(* IEC 61131-3 sources: Zbiorniki_user/Temp/Import/MpRecipe, 4 files *)

(* ---- MpRecipe.typ ---- *)
TYPE
	MpRecipeStatusIDType : 	STRUCT
		ID : MpRecipeErrorEnum; (*Error code for mapp component*)
		Severity : MpComSeveritiesEnum; (*Describes the type of information supplied by the status ID (success, information, warning, error)*)
		Code : UINT; (*Code for the status ID. This error number can be used to search for additional information in the help system*)
	END_STRUCT;
	MpRecipeDiagType : 	STRUCT
		StatusID : MpRecipeStatusIDType; (*StatusID diagnostics structure*)
	END_STRUCT;
	MpRecipeInfoType : 	STRUCT
		Diag : MpRecipeDiagType; (*Diagnostic structure for the status ID*)
	END_STRUCT;
	MpRecipeUISetupConfirmType : 	STRUCT
		RecipeLoad : BOOL; (*Enables a confirmation window when loading a recipe*)
		RecipeSave : BOOL; (*Enables a confirmation window when saving a recipe*)
		RecipeCreate : BOOL; (*Enables a confirmation window when creating a recipe	*)
		RecipeDelete : BOOL; (*Enables a confirmation window when creating a recipe*)
		RecipeRename : BOOL; (*Enables a confirmation window when renaming a recipe*)
	END_STRUCT;
	MpRecipeUISetupType : 	STRUCT
		RecipeListSize : UINT := 20; (*Number of recipes to be displayed on one page of the list in the HMI application*)
		RecipeListScrollWindow : USINT := 1; (*Determines how many entries from the list are displayed in advance when scrolling up and down*)
		Confirmation : MpRecipeUISetupConfirmType; (*Displaying the confirmation window*)
		AutoLoadHeader : BOOL; (*Header info of a recipe should be loaded automatically when a recipe is selected (like a preview) *)
	END_STRUCT;
	MpRecipeUIMessageEnum :
		(
		mpRECIPE_UI_MSG_NONE := 0, (*No dialog is required*)
		mpRECIPE_UI_MSG_CONFIRM_LOAD := 1, (*Dialog box for confirming the loading procedure*)
		mpRECIPE_UI_MSG_CONFIRM_SAVE := 2, (*Dialog box for confirming the saving procedure*)
		mpRECIPE_UI_MSG_CONFIRM_CREATE := 3, (*Dialog box for confirming the creation of a new recipe	*)
		mpRECIPE_UI_MSG_CONFIRM_DELETE := 4, (*Dialog box for confirming the deletion of an existing recipe*)
		mpRECIPE_UI_MSG_CONFIRM_RENAME := 5 (*Dialog box for confirming the renaming of an existing recipe*)
		);
	MpRecipeUIStatusEnum :
		(
		mpRECIPE_UI_STATUS_IDLE := 0, (*Indicates that no process is currently active*)
		mpRECIPE_UI_STATUS_LOAD := 1, (*A recipe is being loaded*)
		mpRECIPE_UI_STATUS_SAVE := 2, (*A recipe is being saved*)
		mpRECIPE_UI_STATUS_CREATE := 3, (*A recipe is being created*)
		mpRECIPE_UI_STATUS_REFRESH := 4, (*The recipe list is being refreshed*)
		mpRECIPE_UI_STATUS_NOTIFY := 5, (*mapp components are being informed that new parameters are to be used*)
		mpRECIPE_UI_STATUS_DELETE := 6, (*A recipe is being deleted*)
		mpRECIPE_UI_STATUS_RENAME := 7, (*A recipe is being renamed*)
		mpRECIPE_UI_STATUS_ERROR := 99 (*The last operation generated an error*)
		);
	MpRecipeUIMessageBoxType : 	STRUCT
		LayerStatus : UINT; (*Visibility of the dialog box *)
		Type : MpRecipeUIMessageEnum; (*Type of dialog box*)
		Confirm : BOOL; (*Confirms the operation*)
		Cancel : BOOL; (*Cancels the operation*)
	END_STRUCT;
	MpRecipeUINewType : 	STRUCT
		FileName : STRING[255]; (*Name of the new recipe*)
		Create : BOOL; (*Creates a new recipe*)
	END_STRUCT;
	MpRecipeUIConnectType : 	STRUCT
		Status : MpRecipeUIStatusEnum; (*Current operation*)
		Recipe : MpRecipeUIRecipeType; (*Access to existing recipes*)
		New : MpRecipeUINewType; (*To create new recipes*)
		MessageBox : MpRecipeUIMessageBoxType; (*Controls dialog boxes*)
		DefaultLayerStatus : UINT; (*Status data point for the default layer of the visualization page where the recipe management system is being displayed*)
	END_STRUCT;
	MpRecipeUIRecipeListType : 	STRUCT
		Names : ARRAY[0..19] OF STRING[255]; (*List of all available recipes (filenames)*)
		SelectedIndex : UINT; (*Index of the entry currently selected in the list*)
		MaxSelection : UINT; (*Index of the last entry in the list*)
		PageUp : BOOL; (*Jumps to the start of the current page and then scrolls up one page at a time *)
		PageDown : BOOL; (*Jumps to the end of the current page and then scrolls down one page at a time *)
		StepUp : BOOL; (*Selects the previous entry in the list*)
		StepDown : BOOL; (*Selects the next entry in the list*)
		RangeStart : REAL; (*Shows a bar indicating which part of the list is currently being displayed-Start [%]*)
		RangeEnd : REAL; (*Shows a bar indicating which part of the list is currently being displayed-End [%]*)
		Sizes : ARRAY[0..19]OF UDINT; (*List of all recipe file sizes*)
		LastModified : ARRAY[0..19]OF STRING[50]; (*List of the last modification dates for all recipe files*)
	END_STRUCT;
	MpRecipeUIHeaderType : 	STRUCT
		Name : STRING[100]; (*Name of the recipe*)
		Description : STRING[255]; (*Comment that describes the recipe*)
		Version : STRING[20]; (*Version of the recipe*)
		DateTime : DATE_AND_TIME; (*Date and time the recipe was created*)
	END_STRUCT;
	MpRecipeUIRecipeType : 	STRUCT
		List : MpRecipeUIRecipeListType; (*List of all available recipes (filenames)*)
		Load : BOOL; (*Loads the selected recipe*)
		Save : BOOL; (*Saves the selected recipe*)
		Filter : STRING[255]; (*Filter used to sort the recipes*)
		SortOrder : MpRecipeUISortOrderEnum; (*Sorts the recipe list*)
		Refresh : BOOL; (*Updates the recipe list*)
		UpdateNotification : BOOL; (*Request to all mapp components to enter the current values of the recipe parameters*)
		Delete : BOOL; (*Deletes the selected recipe*)
		Rename : BOOL; (*Renames the currently selected recipe*)
		NewFileName : STRING[255]; (*Name of the new recipe*)
		Header : MpRecipeUIHeaderType; (*The header info of the currently selected recipe (is only loaded if the option is enabled in UISetup)*)
	END_STRUCT;
	MpRecipeXmlInfoType : 	STRUCT
		FileSize : UDINT; (*Size of the recipe stored on the respective data storage medium*)
		PendingSync : UDINT; (*Number of pending save notifications ("SaveNotification") that have not yet been confirmed*)
		Diag : MpRecipeDiagType; (*Diagnostic structure for the status ID *)
		LastLoadedRecipe : STRING[255]; (*The name of the last loaded recipe*)
	END_STRUCT;
	MpRecipeUISortOrderEnum :
		(
		mpRECIPE_UI_SORT_ASCENDING := 0, (*Sorts in ascending (alphabetic) order*)
		mpRECIPE_UI_SORT_DESCENDING := 1, (*Sorts in descending (alphabetic) order*)
		mpRECIPE_UI_SORT_DATE_ASCENDING := 2, (*Sorts in ascending (date/time) order*)
		mpRECIPE_UI_SORT_DATE_DESCENDING := 3 (*Sorts in descending (date/time) order*)
		);
	MpRecipeXmlHeaderType : 	STRUCT
		Name : STRING[100]; (*Name of the recipe*)
		Description : STRING[255]; (*Comment that describes the recipe*)
		Version : STRING[20]; (*Version of the recipe*)
		DateTime : DATE_AND_TIME; (*Date and time the recipe was created*)
	END_STRUCT;
	MpRecipeXmlLoadEnum :
		(
		mpRECIPE_XML_LOAD_ALL := 0, (*Loads the entire content of the recipe*)
		mpRECIPE_XML_LOAD_HEADER := 1 (*Loads only the recipe's header*)
		);
	MpRecipeCsvHeaderType : 	STRUCT
		Name : STRING[100]; (*Name of the recipe*)
		Description : STRING[255]; (*Comment that describes the recipe*)
		Version : STRING[20]; (*Version of the recipe*)
		DateTime : DATE_AND_TIME; (*Date and time the recipe was created*)
	END_STRUCT;
	MpRecipeCsvInfoType : 	STRUCT
		FileSize : UDINT; (*Size of the recipe stored on the respective data storage medium*)
		PendingSync : UDINT; (*Number of pending save notifications ("SaveNotification") that have not yet been confirmed*)
		LastLoadedRecipe : STRING[255]; (*The name of the last loaded recipe*)
		Diag : MpRecipeDiagType; (*Diagnostic structure for the status ID *)
	END_STRUCT;
	MpRecipeCsvLoadEnum :
		(
		mpRECIPE_CSV_LOAD_ALL := 0, (*Loads the entire content of the recipe*)
		mpRECIPE_CSV_LOAD_HEADER := 1 (*Loads only the recipe's header*)
		);
END_TYPE

(* ---- MpRecipeAlarm.typ ---- *)
TYPE
    MpRecipeXmlAlarmEnum :
        ( (* Alarms of MpRecipe Xml *)
        mpRECIPE_ALM_SAVE_FAILED := 0, (* Saving of recipe failed. *)
        mpRECIPE_ALM_SAVE_FAILED_PART := 1, (* Saving of recipe failed partially. Parts of the recipe could be saved. *)
        mpRECIPE_ALM_LOAD_FAILED := 2, (* Loading of recipe failed. *)
        mpRECIPE_ALM_LOAD_FAILED_PART := 3 (* Loading of recipe failed partially. Parts of the recipe could be loaded. *)
    );
END_TYPE

(* ---- MpRecipeError.typ ---- *)
TYPE
    MpRecipeErrorEnum :
        ( (* Error numbers of library MpRecipe *)
        mpRECIPE_NO_ERROR := 0, (* No error *)
        mpRECIPE_ERR_ACTIVATION := -1064239103, (* Could not create component [Error: 1, 0xc0910001] *)
        mpRECIPE_ERR_MPLINK_NULL := -1064239102, (* MpLink is NULL pointer [Error: 2, 0xc0910002] *)
        mpRECIPE_ERR_MPLINK_INVALID := -1064239101, (* MpLink connection not allowed [Error: 3, 0xc0910003] *)
        mpRECIPE_ERR_MPLINK_CHANGED := -1064239100, (* MpLink modified [Error: 4, 0xc0910004] *)
        mpRECIPE_ERR_MPLINK_CORRUPT := -1064239099, (* Invalid MpLink contents [Error: 5, 0xc0910005] *)
        mpRECIPE_ERR_MPLINK_IN_USE := -1064239098, (* MpLink already in use [Error: 6, 0xc0910006] *)
        mpRECIPE_ERR_CONFIG_INVALID := -1064239091, (* Invalid Configuration [Error: 13, 0xc091000d] *)
        mpRECIPE_ERR_SAVE_DATA := -1064140799, (* Failed to create recipe file {2:File} using device {3:Device} (Error cause: {1:ErrorNumber}) [Error: 32769, 0xc0928001] *)
        mpRECIPE_ERR_LOAD_DATA := -1064140798, (* Failed to load recipe from {2:File} using device {3:Device} (Error cause: {1:ErrorNumber}) [Error: 32770, 0xc0928002] *)
        mpRECIPE_ERR_INVALID_FILE_DEV := -1064140797, (* Invalid file device [Error: 32771, 0xc0928003] *)
        mpRECIPE_ERR_INVALID_FILE_NAME := -1064140796, (* Invalid filename [Error: 32772, 0xc0928004] *)
        mpRECIPE_ERR_CMD_IN_PROGRESS := -1064140795, (* Component currently executing command [Error: 32773, 0xc0928005] *)
        mpRECIPE_WRN_SAVE_WITH_WARN := -2137882618, (* Warnings while saving recipe [Warning: 32774, 0x80928006] *)
        mpRECIPE_WRN_LOAD_WITH_WARN := -2137882617, (* Warnings while loading recipe [Warning: 32775, 0x80928007] *)
        mpRECIPE_ERR_SAVE_WITH_ERRORS := -1064140792, (* Failed to write to recipe file {2:File} (Error cause: {1:ErrorNumber}) [Error: 32776, 0xc0928008] *)
        mpRECIPE_ERR_LOAD_WITH_ERRORS := -1064140791, (* Error converting recipe to parameters [Error: 32777, 0xc0928009] *)
        mpRECIPE_ERR_MISSING_RECIPE := -1064140790, (* No connection to parent component [Error: 32778, 0xc092800a] *)
        mpRECIPE_ERR_MISSING_MPFILE := -1064140789, (* No connection to file manager [Error: 32779, 0xc092800b] *)
        mpRECIPE_ERR_INVALID_SORT_ORDER := -1064140788, (* Invalid sort order selected [Error: 32780, 0xc092800c] *)
        mpRECIPE_WRN_MISSING_UICONNECT := -2137882611, (* Invalid value for "UIConnect" [Warning: 32781, 0x8092800d] *)
        mpRECIPE_ERR_INVALID_PV_NAME := -1064140786, (* Invalid PV [Error: 32782, 0xc092800e] *)
        mpRECIPE_ERR_INVALID_LOAD_TYPE := -1064140785, (* Invalid LoadType [Error: 32783, 0xc092800f] *)
        mpRECIPE_ERR_LISTING_FILES := -1064140784, (* Error creating file list [Error: 32784, 0xc0928010] *)
        mpRECIPE_ERR_PV_NAME_NULL := -1064140783, (* PV name is NULL [Error: 32785, 0xc0928011] *)
        mpRECIPE_WRN_NO_PV_REGISTERED := -2137882606, (* No PV registered [Warning: 32786, 0x80928012] *)
        mpRECIPE_ERR_SYNC_SAVE_ACTIVE := -1064140781, (* Saving active [Error: 32787, 0xc0928013] *)
        mpRECIPE_ERR_DELETING_FILE := -1064140780, (* Failed to delete recipe {2:Recipe} from device {3:Device} (Error cause: {1:ErrorNumber}) [Error: 32788, 0xc0928014] *)
        mpRECIPE_WRN_EMPTY_RECIPE := -2137882603, (* Saving empty recipe file [Warning: 32789, 0x80928015] *)
        mpRECIPE_INF_WAIT_RECIPE_FB := 1083342870, (* Waiting for parent recipe component [Informational: 32790, 0x40928016] *)
        mpRECIPE_ERR_RENAMING_FILE := -1064140777, (* Failed to rename recipe {2:FromName} to {3:ToName} (Error cause: {1:ErrorNumber} [Error: 32791, 0xc0928017] *)
        mpRECIPE_WRN_NO_PV_FOUND := -2137882600, (* None of the registered PVs were found in the recipe file while loading. The file might be corrupted. [Warning: 32792, 0x80928018] *)
        mpRECIPE_WRN_LIST_SIZE := -2137882599 (* The UISetup.RecipeListSize {2:Size} is out of limit (1-20). [Warning: 32793, 0x80928019] *)
        );
END_TYPE

(* ---- MpRecipe.fun ---- *)
FUNCTION_BLOCK MpRecipeRegParSync (*Declare a PV as a recipe parameter and perform synchronisation*) (* $GROUP=mapp Services,$CAT=XML Recipe,$GROUPICON=Icon_mapp.png,$CATICON=Icon_MpRecipe.png *)
	VAR_INPUT
		MpLink : REFERENCE TO MpComIdentType; (*Connection to mapp*) (* *) (*#PAR#;*)
		Enable : BOOL; (*Enables/Disables the function block *) (* *) (*#PAR#;*)
		ErrorReset : BOOL; (*Resets function block errors*) (* *) (*#PAR#;*)
		PVName : REFERENCE TO STRING[100]; (*Name of the PV that should be saved to the recipe*) (* *) (*#PAR#;*)
		Category : REFERENCE TO STRING[50]; (*Name of the category used to organize the parameters*) (* *) (*#PAR#OPT#;*)
		ConfirmSave : BOOL; (*Confirms that the current data of the registered PV can be saved to the recipe. This is used in connection with "SaveNotification"*) (* *) (*#CMD#;*)
	END_VAR
	VAR_OUTPUT
		Active : BOOL; (*Indicates whether the function block is active*) (* *) (*#PAR#;*)
		Error : BOOL; (*Indicates that the function block is in an error state or a command was not executed correctly*) (* *) (*#PAR#;*)
		StatusID : DINT; (*Status information about the function block*) (* *) (*#PAR#; *)
		UpdateNotification : BOOL; (*TRUE if a new recipe has been loaded and the registered PV contains new values. This is automatically reset after one cycle*) (* *) (*#CMD#OPT#;*)
		SaveNotification : BOOL; (*TRUE if a recipe is saved and new data should be copied to the recipe, but before the data is actually transferred to the recipe. This is used in connection with "ConfirmSave"*) (* *) (*#CMD#;*)
		Info : MpRecipeInfoType; (*Additional information about the component*) (* *) (*#CMD#;*)
	END_VAR
	VAR
		Internal : {REDUND_UNREPLICABLE} MpComInternalDataType; (*Internal stucture*) (* *) (*#OMIT#;*)
	END_VAR
END_FUNCTION_BLOCK

FUNCTION_BLOCK MpRecipeRegPar (*Declare a PV as a recipe parameter*) (* $GROUP=mapp Services,$CAT=XML Recipe,$GROUPICON=Icon_mapp.png,$CATICON=Icon_MpRecipe.png *)
	VAR_INPUT
		MpLink : REFERENCE TO MpComIdentType; (* Connection to mapp*) (* *) (*#PAR#;*)
		Enable : BOOL; (*Enables/Disables the function block*) (* *) (*#PAR#;*)
		ErrorReset : BOOL; (*Resets function block errors*) (* *) (*#PAR#;*)
		PVName : REFERENCE TO STRING[100]; (*Name of the PV that should be saved to the recipe*) (* *) (*#PAR#;*)
		Category : REFERENCE TO STRING[50]; (*Name of the category used to organize the parameters*) (* *) (*#PAR#OPT#;*)
	END_VAR
	VAR_OUTPUT
		Active : BOOL; (*Indicates whether the function block is active*) (* *) (*#PAR#;*)
		Error : BOOL; (*Indicates that the function block is in an error state or a command was not executed correctly*) (* *) (*#PAR#;*)
		StatusID : DINT; (*Status information about the function block*) (* *) (*#PAR#; *)
		UpdateNotification : BOOL; (*TRUE if a new recipe has been loaded and the registered PV contains new values. This is automatically reset after one cycle*) (* *) (*#CMD#OPT#;*)
		Info : MpRecipeInfoType; (*Additional information about the component*) (* *) (*#CMD#;*)
	END_VAR
	VAR
		Internal : {REDUND_UNREPLICABLE} MpComInternalDataType; (*Internal stucture*) (* *) (*#OMIT#;*)
	END_VAR
END_FUNCTION_BLOCK

FUNCTION_BLOCK MpRecipeXml (*Load/save parameters from/to an XML file*) (* $GROUP=mapp Services,$CAT=XML Recipe,$GROUPICON=Icon_mapp.png,$CATICON=Icon_MpRecipe.png *)
	VAR_INPUT
		MpLink : REFERENCE TO MpComIdentType; (*Connection to mapp*) (* *) (*#PAR#;*)
		Enable : BOOL; (*Enables/Disables the function block*) (* *) (*#PAR#;*)
		ErrorReset : BOOL; (*Resets function block errors*) (* *) (*#PAR#;*)
		DeviceName : REFERENCE TO STRING[50]; (*File device (data storage medium) where the files are stored*) (* *) (*#CMD#;*)
		FileName : REFERENCE TO STRING[255]; (*Name of the file that contains the recipe*) (* *) (*#CMD#;*)
		Header : REFERENCE TO MpRecipeXmlHeaderType; (*Header information that is either written or read*) (* *) (*#CMD#OPT#;*)
		Category : REFERENCE TO STRING[50]; (*Name of the category used to organize the parameters*) (* *) (*#CMD#OPT#;*)
		LoadType : MpRecipeXmlLoadEnum; (*Defines how the recipe is loaded. By default, the entire recipe is loaded*) (* *) (*#CMD#OPT#;*)
		Load : BOOL; (*Loads the recipe parameters from the specified file ("FileName")*) (* *) (*#CMD#;*)
		Save : BOOL; (*Saves the current recipe parameters to a defined file*) (* *) (*#CMD#;*)
		UpdateNotification : BOOL; (*A rising edge on this input induces all MpRecipeRegPar and MpRecipeRegParSync instances to provide information about new recipe values on their "UpdateNotification" output for one cycle*) (* *) (*#CMD#OPT#;*)
	END_VAR
	VAR_OUTPUT
		Active : BOOL; (*Indicates whether the function block is active*) (* *) (*#PAR#;*)
		Error : BOOL; (*Indicates that the function block is in an error state or a command was not executed correctly*) (* *) (*#PAR#;*)
		StatusID : DINT; (*Status information about the function block*) (* *) (*#PAR#; *)
		CommandBusy : BOOL; (*Function block currently executing command*) (* *) (*#CMD#OPT#;*)
		CommandDone : BOOL; (*Command successfully executed by function block*) (* *) (*#CMD#;*)
		Info : MpRecipeXmlInfoType; (*Additional information about the component*) (* *) (*#CMD#;*)
	END_VAR
	VAR
		Internal : {REDUND_UNREPLICABLE} MpComInternalDataType; (*Internal stucture*) (* *) (*#OMIT#;*)
	END_VAR
END_FUNCTION_BLOCK

FUNCTION_BLOCK MpRecipeUI (*UI connection to a VC4 recipe page*) (* $GROUP=mapp Services,$CAT=XML Recipe,$GROUPICON=Icon_mapp.png,$CATICON=Icon_MpRecipe.png *)
	VAR_INPUT
		MpLink : REFERENCE TO MpComIdentType; (*Connection to mapp*) (* *) (*#PAR#;*)
		Enable : BOOL; (*Enables/Disables the function block*) (* *) (*#PAR#;*)
		ErrorReset : BOOL; (*Resets function block errors*) (* *) (*#PAR#;*)
		UISetup : {REDUND_UNREPLICABLE} MpRecipeUISetupType; (*Used to configure the elements connected to the HMI application*) (* *) (*#PAR#;*)
		UIConnect : REFERENCE TO MpRecipeUIConnectType; (*This structure contains the parameters needed for the connection to the HMI application*) (* *) (*#CMD#;*)
	END_VAR
	VAR_OUTPUT
		Active : BOOL; (*Indicates whether the function block is active*) (* *) (*#PAR#;*)
		Error : BOOL; (*Indicates that the function block is in an error state or a command was not executed correctly*) (* *) (*#PAR#;*)
		StatusID : DINT; (*Status information about the function block*) (* *) (*#PAR#;*)
		Info : MpRecipeInfoType; (*Additional information about the component*) (* *) (*#CMD;*)
	END_VAR
	VAR
		Internal : {REDUND_UNREPLICABLE} MpComInternalDataType; (*Internal stucture*) (* *) (*#OMIT#;*)
	END_VAR
END_FUNCTION_BLOCK

FUNCTION_BLOCK MpRecipeCsv (*Load/save parameters from/to an CSV file*) (* $GROUP=mapp Services,$CAT=CSV Recipe,$GROUPICON=Icon_mapp.png,$CATICON=Icon_MpRecipe.png *)
	VAR_INPUT
		MpLink : REFERENCE TO MpComIdentType; (*Connection to mapp*) (* *) (*#PAR#;*)
		Enable : BOOL; (*Enables/Disables the function block*) (* *) (*#PAR#;*)
		ErrorReset : BOOL; (*Resets function block errors*) (* *) (*#PAR#;*)
		DeviceName : REFERENCE TO STRING[50]; (*File device (data storage medium) where the files are stored*) (* *) (*#CMD#;*)
		FileName : REFERENCE TO STRING[255]; (*Name of the file that contains the recipe*) (* *) (*#CMD#;*)
		Header : REFERENCE TO MpRecipeCsvHeaderType; (*Header information that is either written or read*) (* *) (*#CMD#OPT#;*)
		Category : REFERENCE TO STRING[50]; (*Name of the category used to organize the parameters*) (* *) (*#CMD#OPT#;*)
		LoadType : MpRecipeCsvLoadEnum; (*Defines how the recipe is loaded. By default, the entire recipe is loaded*) (* *) (*#CMD#OPT#;*)
		Load : BOOL; (*Loads the recipe parameters from the specified file ("FileName")*) (* *) (*#CMD#;*)
		Save : BOOL; (*Saves the current recipe parameters to a defined file*) (* *) (*#CMD#;*)
		UpdateNotification : BOOL; (*A rising edge on this input induces all MpRecipeRegPar and MpRecipeRegParSync instances to provide information about new recipe values on their "UpdateNotification" output for one cycle*) (* *) (*#CMD#OPT#;*)
	END_VAR
	VAR_OUTPUT
		Active : BOOL; (*Indicates whether the function block is active*) (* *) (*#PAR#;*)
		Error : BOOL; (*Indicates that the function block is in an error state or a command was not executed correctly*) (* *) (*#PAR#;*)
		StatusID : DINT; (*Status information about the function block*) (* *) (*#PAR#; *)
		CommandBusy : BOOL; (*Function block currently executing command*) (* *) (*#CMD#OPT#;*)
		CommandDone : BOOL; (*Command successfully executed by function block*) (* *) (*#CMD#;*)
		Info : MpRecipeCsvInfoType; (*Additional information about the component*) (* *) (*#CMD#;*)
	END_VAR
	VAR
		Internal : {REDUND_UNREPLICABLE} MpComInternalDataType; (*Internal stucture*) (* *) (*#OMIT#;*)
	END_VAR
END_FUNCTION_BLOCK
